(* IEC 61131-3 sources: llm-plc-st-eval/data/processed_v2_primera/gpt-4o/B5/few_shot, 3 files *)

(* ---- ejec_1.st ---- *)
FUNCTION_BLOCK FB_Ventilador
VAR_INPUT
    quemadorOn : BOOL; (* Estado del quemador *)
END_VAR
VAR_OUTPUT
    ventilador : BOOL; (* Estado del ventilador *)
END_VAR
VAR
    tRetraso : TON; (* Temporizador de retardo *)
END_VAR

(* El ventilador funciona mientras el quemador está encendido o durante 30 segundos adicionales después de apagarse *)
tRetraso(IN := NOT quemadorOn, PT := T#30S);
ventilador := quemadorOn OR tRetraso.Q;
END_FUNCTION_BLOCK

(* ---- ejec_2.st ---- *)
FUNCTION_BLOCK FB_Ventilador
VAR_INPUT
    quemadorOn : BOOL; (* Estado del quemador *)
END_VAR
VAR_OUTPUT
    ventilador : BOOL; (* Estado del ventilador *)
END_VAR
VAR
    tRetraso : TON; (* Temporizador de retardo *)
END_VAR

(* El ventilador funciona mientras el quemador está encendido o durante 30 segundos adicionales después de apagarse *)
tRetraso(IN := NOT quemadorOn, PT := T#30S);
ventilador := quemadorOn OR tRetraso.Q;
END_FUNCTION_BLOCK

(* ---- ejec_3.st ---- *)
FUNCTION_BLOCK FB_Ventilador
VAR_INPUT
    quemadorOn : BOOL; (* Estado del quemador *)
END_VAR
VAR_OUTPUT
    ventilador : BOOL; (* Estado del ventilador *)
END_VAR
VAR
    tRetraso : TON; (* Temporizador de retardo *)
END_VAR

(* El ventilador funciona mientras el quemador está encendido o durante 30 segundos después de apagarse *)
tRetraso(IN := NOT quemadorOn, PT := T#30S);
ventilador := quemadorOn OR tRetraso.Q;
END_FUNCTION_BLOCK
